FUNCTION_BLOCK AUTO_RESTART (* Migrated from IEC 61131-3 ST *)
  (* Standard: 61499-2 *)
  (* Version 1.0, 2026-11-06, st2fb *)
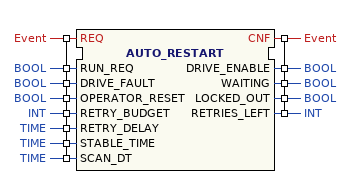
  EVENT_INPUT
    REQ WITH RUN_REQ, DRIVE_FAULT, OPERATOR_RESET, RETRY_BUDGET, RETRY_DELAY, STABLE_TIME, SCAN_DT;
  END_EVENT
  EVENT_OUTPUT
    CNF WITH DRIVE_ENABLE, WAITING, LOCKED_OUT, RETRIES_LEFT;
  END_EVENT
  VAR_INPUT
    RUN_REQ : BOOL;
    DRIVE_FAULT : BOOL;
    OPERATOR_RESET : BOOL;
    RETRY_BUDGET : INT;
    RETRY_DELAY : TIME;
    STABLE_TIME : TIME;
    SCAN_DT : TIME;
  END_VAR
  VAR_OUTPUT
    DRIVE_ENABLE : BOOL;
    WAITING : BOOL;
    LOCKED_OUT : BOOL;
    RETRIES_LEFT : INT;
  END_VAR
  VAR
    ST2FB_NOW : TIME := T#0s;
    FAULT_EDGE_CLK : BOOL;
    FAULT_EDGE_Q : BOOL;
    FAULT_EDGE_M : BOOL;
    BUDGET_CD : BOOL;
    BUDGET_LD : BOOL;
    BUDGET_PV : INT;
    BUDGET_Q : BOOL;
    BUDGET_CV : INT;
    BUDGET_CD_T_Q : BOOL;
    BUDGET_CD_T_M : BOOL;
    LOCKOUT_S : BOOL;
    LOCKOUT_R1 : BOOL;
    LOCKOUT_Q1 : BOOL;
    WAIT_TIMER_IN : BOOL;
    WAIT_TIMER_PT : TIME;
    WAIT_TIMER_Q : BOOL;
    WAIT_TIMER_ET : TIME;
    WAIT_TIMER_STATE : INT;
    WAIT_TIMER_PREV_IN : BOOL;
    WAIT_TIMER_START_TIME : TIME;
    STABLE_TIMER_IN : BOOL;
    STABLE_TIMER_PT : TIME;
    STABLE_TIMER_Q : BOOL;
    STABLE_TIMER_ET : TIME;
    STABLE_TIMER_STATE : INT;
    STABLE_TIMER_PREV_IN : BOOL;
    STABLE_TIMER_START_TIME : TIME;
    LOADED : BOOL;
  END_VAR
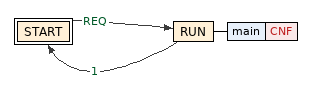
  EC_STATES
    START;
    RUN : main -> CNF;
  END_STATES
  EC_TRANSITIONS
    START TO RUN := REQ;
    RUN TO START := 1;
  END_TRANSITIONS
  ALGORITHM main IN ST:
ST2FB_NOW := ST2FB_NOW + SCAN_DT;

FAULT_EDGE_CLK := DRIVE_FAULT;
FAULT_EDGE_Q := FAULT_EDGE_CLK AND NOT FAULT_EDGE_M;
FAULT_EDGE_M := FAULT_EDGE_CLK;

STABLE_TIMER_IN := DRIVE_ENABLE AND NOT DRIVE_FAULT;
STABLE_TIMER_PT := STABLE_TIME;
IF (STABLE_TIMER_STATE = 0) AND NOT STABLE_TIMER_PREV_IN AND STABLE_TIMER_IN THEN
  STABLE_TIMER_STATE := 1;
  STABLE_TIMER_Q := FALSE;
  STABLE_TIMER_START_TIME := ST2FB_NOW;
ELSE
  IF NOT STABLE_TIMER_IN THEN
    STABLE_TIMER_ET := T#0s;
    STABLE_TIMER_Q := FALSE;
    STABLE_TIMER_STATE := 0;
  ELSIF STABLE_TIMER_STATE = 1 THEN
    IF STABLE_TIMER_START_TIME + STABLE_TIMER_PT <= ST2FB_NOW THEN
      STABLE_TIMER_STATE := 2;
      STABLE_TIMER_Q := TRUE;
      STABLE_TIMER_ET := STABLE_TIMER_PT;
    ELSE
      STABLE_TIMER_ET := ST2FB_NOW - STABLE_TIMER_START_TIME;
    END_IF;
  END_IF;
END_IF;
STABLE_TIMER_PREV_IN := STABLE_TIMER_IN;

BUDGET_CD := FAULT_EDGE_Q;
BUDGET_LD := NOT LOADED OR OPERATOR_RESET OR STABLE_TIMER_Q;
BUDGET_PV := RETRY_BUDGET;
BUDGET_CD_T_Q := BUDGET_CD AND NOT BUDGET_CD_T_M;
BUDGET_CD_T_M := BUDGET_CD;
IF BUDGET_LD THEN
  BUDGET_CV := BUDGET_PV;
ELSIF BUDGET_CD_T_Q AND (BUDGET_CV > 0) THEN
  BUDGET_CV := BUDGET_CV - 1;
END_IF;
BUDGET_Q := BUDGET_CV <= 0;

LOADED := TRUE;
RETRIES_LEFT := BUDGET_CV;

LOCKOUT_S := FAULT_EDGE_Q AND BUDGET_Q;
LOCKOUT_R1 := OPERATOR_RESET;
LOCKOUT_Q1 := NOT LOCKOUT_R1 AND (LOCKOUT_S OR LOCKOUT_Q1);
LOCKED_OUT := LOCKOUT_Q1;

IF DRIVE_FAULT THEN
  WAITING := TRUE;
END_IF;

WAIT_TIMER_IN := WAITING AND NOT DRIVE_FAULT;
WAIT_TIMER_PT := RETRY_DELAY;
IF (WAIT_TIMER_STATE = 0) AND NOT WAIT_TIMER_PREV_IN AND WAIT_TIMER_IN THEN
  WAIT_TIMER_STATE := 1;
  WAIT_TIMER_Q := FALSE;
  WAIT_TIMER_START_TIME := ST2FB_NOW;
ELSE
  IF NOT WAIT_TIMER_IN THEN
    WAIT_TIMER_ET := T#0s;
    WAIT_TIMER_Q := FALSE;
    WAIT_TIMER_STATE := 0;
  ELSIF WAIT_TIMER_STATE = 1 THEN
    IF WAIT_TIMER_START_TIME + WAIT_TIMER_PT <= ST2FB_NOW THEN
      WAIT_TIMER_STATE := 2;
      WAIT_TIMER_Q := TRUE;
      WAIT_TIMER_ET := WAIT_TIMER_PT;
    ELSE
      WAIT_TIMER_ET := ST2FB_NOW - WAIT_TIMER_START_TIME;
    END_IF;
  END_IF;
END_IF;
WAIT_TIMER_PREV_IN := WAIT_TIMER_IN;

IF WAIT_TIMER_Q OR NOT RUN_REQ THEN
  WAITING := FALSE;
END_IF;
DRIVE_ENABLE := RUN_REQ AND NOT DRIVE_FAULT AND NOT WAITING AND NOT LOCKED_OUT;
  END_ALGORITHM
END_FUNCTION_BLOCK
